// TIA Portal V21 export
// export: Created 2026-11-10T07:35:10.6923853Z, ExportSetting WithDefaults, DisplayName Totally Integrated Automation Portal, DisplayVersion V21 Update 3, DisplayName STEP 7 Professional, DisplayVersion V21 Update 3, DisplayName STEP 7 Safety, DisplayVersion V21, DisplayName Tech WebApplication, DisplayVersion V21, DisplayName WinCC Basic/Comfort/Advanced, DisplayVersion V21 Update 3, DisplayName WinCC Unified, DisplayVersion V21 Update 3
FUNCTION_BLOCK "FB_Lad_ex098"   // FB70, LAD
{ S7_Optimized_Access := 'TRUE' }
VERSION : 0.1
// stored: AutoNumber true, IsIECCheckEnabled false, IsRetainMemResEnabled false, MemoryReserve 100, SetENOAutomatically false, UDAEnableTagReadback false
   VAR_INPUT
      v_ioid : Byte;
      v_laddr : HW_IO;
      v_recnum : Byte;
      v_ret_val : Int;
   END_VAR
   VAR_IN_OUT
      v_record : Variant;
   END_VAR
BEGIN

REGION Network 1: RD_DPARM - Read data record from configured system data
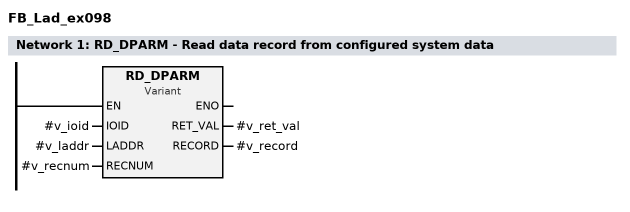
   RUNG wire#powerrail
      { S7_Templates := "[record_type := Variant, laddr_type := HW_IO]" } RD_DPARM(IOID := #v_ioid, LADDR := #v_laddr, RECNUM := #v_recnum, RET_VAL => #v_ret_val, RECORD => #v_record)
   END_RUNG
   // the same network as SCL:
   #v_ret_val := RD_DPARM(IOID := #v_ioid, LADDR := #v_laddr, RECNUM := #v_recnum, RECORD => #v_record);
END_REGION
END_FUNCTION_BLOCK
